(* Communication structure from drive to plc *)

TYPE ST_FORCETOPLC :
STRUCT

END_STRUCT
END_TYPE

(* stored: Version 1.1.0.1, ProductVersion 3.1.4024.15
   DUT ST_FORCETOPLC: Id {31c28a24-7b24-492c-a3e6-c85a430ee6f9} *)
